Staubli VAL3: HMI_safepoint.pjx

--- HMI_safepoint.pjx ---
Parameters version=s8.12.1Cs9_BS2449 stackSize=5000 millimeterUnit=true
Program file=bind.pgx
Program file=main.pgx
Program file=movePoint.pgx
Program file=onStart.pgx
Program file=setActive.pgx
Program file=showActive.pgx
Program file=showCoord.pgx
Program file=start.pgx
Program file=stop.pgx
Program file=teachPoint.pgx
Data file=HMI_safepoint.dtx
Library alias=util path=Disk://HMI_cs9/HMI_util/HMI_util.pjx
Library alias=safeTemp path=Disk://data/CustomerLib/default/safeData/safeData.pjx
Library alias=rs path=Disk://source/projectSource/robotStatus/robotStatus.pjx
Library alias=savedata path=Disk://source/saveData/saveData.pjx
Library alias=saveData path=Disk://source/saveData/saveData.pjx

--- HMI_safepoint.dtx ---
mdesc mNomSpeed
bool bBack
bool bTeach
bool bMove
string sList
string sSelPoint
bool bActive
string sTRSF[6]
string sLastPoint
mdesc mSimulate = {blend=off}

--- main.pgx ---
public program main()
  local num l_nIndex
  local bool l_bResult
  local bool l_bRefresh
  local bool l_bExit
begin
  do
    if util:sPage!="safepoint"
      util:sPage="safepoint"
      call onStart()
      call bind()
      userPage(util:sPage)
      delay(0.5)
    endIf
    if sLastPoint!=sSelPoint
      sLastPoint=sSelPoint
      toNum(sSelPoint,l_nIndex,l_bResult)
      if l_bResult
        l_bRefresh=true
         call showActive(l_nIndex)
      endIf
    endIf


    if bBack
      bBack=false
      safeTemp:libSave()
      delay(0.1)
      l_bExit=true
    elseIf bTeach
      bTeach=false
      call teachPoint(l_nIndex)
      l_bRefresh=true
    elseIf bMove
      bMove=false
      call movePoint(l_nIndex)
      l_bRefresh=true
    elseIf bActive!= safeTemp:sSPoint[l_nIndex].bActive and sSelPoint!=""
      safeTemp:sSPoint[l_nIndex].bActive=(bActive==true)
      safeTemp:libSave()
      delay(0.1)
    endIf
    if l_bRefresh
      l_bRefresh=false
      call showCoord(l_nIndex)

    endIf

    call util:jogMode(0,0)
    delay(0)
  until l_bExit==true

end

--- start.pgx ---
program start()
begin
  call main()
end

--- bind.pgx ---
program bind()
  local string l_slbl
  local num l_i
begin
  userPageBindClick("safepoint","btnback",bBack,true)
  userPageBindClick("safepoint","btn1",bTeach,true)
  userPageBindClick("safepoint","btn2",bMove,true)

  userPageBind("safepoint","lst1","options",sList,size(sList),"r")
  userPageBind("safepoint","lst1","value",sSelPoint,1,"rw")

  userPageBind("safepoint","chk1","checked",bActive,1,"rw")

  for l_i = 0 to 5
    l_slbl="lbl3"+toString("",l_i)
    userPageBind("safepoint",l_slbl,"innerHTML",sTRSF[l_i],1,"r")
  endFor
end

--- movePoint.pgx ---
program movePoint(num x_nIndex)
  local bool l_bResult
  local jointRx l_joint
begin
  l_bResult=userPageConfirm("是否移动到点位："+toString("",x_nIndex)+"?")
  if l_bResult and rs:_nOmacStat==9
    resetMotion()
    l_bResult=pointToJoint(flange,herej(),safeTemp:sSPoint[x_nIndex].pPointRx,l_joint)
    if l_bResult
      movej(safeTemp:sSPoint[x_nIndex].pPointRx,flange,mSimulate)
    else
      popUpMsg("无法移动到该安全点位")
    endIf
  endIf
  if rs:_nOmacStat!=9
    userPageAlert("机器人当前状态不满足，无法执行移动")
  endIf
end

--- onStart.pgx ---
public program onStart()
  local num l_i
begin
  call saveData:setBaseJOG(saveData:nJogTool)
  resize(sList,1,size(safeTemp:sSPoint))
  for l_i = 0 to size(sList)-1
    sList[l_i]=toString("",l_i)+","+safeTemp:sSPoint[l_i].sName
  endFor

  sSelPoint=""
  sLastPoint=""
  bActive=false

  for l_i = 0 to size(sTRSF)-1
    sTRSF[l_i]=""
  endFor

end

--- setActive.pgx ---
program setActive(num x_nIndex)
begin
  safeTemp:sSPoint[x_nIndex].bActive=(bActive==true)
end

--- showActive.pgx ---
program showActive(num x_nIndex)
begin
  bActive=(safeTemp:sSPoint[x_nIndex].bActive==true)
end

--- showCoord.pgx ---
program showCoord(num x_nIndex)
begin
  sTRSF[0]=toString(".2",safeTemp:sSPoint[x_nIndex].pPointRx.trsf.x)
  sTRSF[1]=toString(".2",safeTemp:sSPoint[x_nIndex].pPointRx.trsf.y)
  sTRSF[2]=toString(".2",safeTemp:sSPoint[x_nIndex].pPointRx.trsf.z)
  sTRSF[3]=toString(".2",safeTemp:sSPoint[x_nIndex].pPointRx.trsf.rx)
  sTRSF[4]=toString(".2",safeTemp:sSPoint[x_nIndex].pPointRx.trsf.ry)
  sTRSF[5]=toString(".2",safeTemp:sSPoint[x_nIndex].pPointRx.trsf.rz)
end

--- stop.pgx ---
program stop()
begin
end

--- teachPoint.pgx ---
program teachPoint(num x_nIndex)
  local bool l_bResult
  local tool l_tTool
begin
  link(l_tTool,flange)
//  call savedata:getTool(1,l_tTool)
  l_bResult=userPageConfirm("是否记录点位："+toString("",x_nIndex)+"?")
  if l_bResult
    safeTemp:sSPoint[x_nIndex].pPointRx=here(flange,world)
    safeTemp:libSave()
    delay(0.1)
  endIf
end
